// TIA Portal V19 export
// export: Created 2026-01-15T10:00:00.0000000Z, ExportSetting WithReadOnly
VAR_GLOBAL   // PLC tag table "Example_Tags"
   Example_Run AT %I0.0 : Bool;   // Run request
   Example_MotorOn AT %Q0.0 : Bool;
   Example_Speed AT %IW64 : Int;
END_VAR
VAR_GLOBAL CONSTANT   // user constants
   Example_MaxSpeed : Int := 1500;
END_VAR
